// TIA Portal V21 export
ORGANIZATION_BLOCK "OB_Cyclic100ms"   // OB35, SCL, CyclicInterrupt
TITLE = Weckalarm 100 ms / Cyclic interrupt 100 ms
{ S7_Optimized_Access := 'TRUE' }
// Ruft FB_SclTimers alle 100 ms mit eigener Instanz auf / Calls FB_SclTimers every 100 ms with its own instance
// stored: AutoNumber false, PhaseOffset 20000, SetENOAutomatically false
   VAR_INPUT
      Initial_Call : Bool;   // Initial call of this OB
      Event_Count : Int;   // Events discarded
   END_VAR
BEGIN

       REGION Timers every 100 ms
           "IDB_SclTimersCyclic"(Start := "LevelHigh", Reset := "StopButton", DelayTime := T#1s);
       END_REGION

       REGION Analyzer C26l
           // The same instance is also called from OB_Main
           "IDB_AnaShared"(Pulse := "LevelHigh");
       END_REGION
END_ORGANIZATION_BLOCK
